(* CODESYS project functionresponse.library
   Company: KOSTAL GmbH & Co.KG
   DocFormat: reStructuredText
   DefaultNamespace: KOSTAL.AF2024.Core.functionResponse
   Version: 1.0.0.0
   Placeholder: KOSTAL.AF2024.Core.functionResponse
   Author: Frank Dümpelmann
   Title: KOSTAL.AF2024.Core.functionResponse

Project tree, tasks and I/O mapping:
  libraries: KOSTAL.AF2024.Core.Settings, * (KOSTAL GmbH & Co.KG); KOSTAL.AF2024.Core.System, * (KOSTAL GmbH & Co.KG)
  DUT/
    interface I_T_functionResponse: CopyTo, status, success
    interface I_T_functionResponse_CopyFrom: CopyFrom
    interface I_T_functionResponse_Owner: clear, CopyFrom, CopyTo, status, success
    function block T_functionResponse [ST]: clear, CopyFrom, CopyTo, status, success
  Project Information/
    function F_GetCompany [ST]
    function F_GetTitle [ST]
    function F_GetVersion [ST]
  Version/
    global variables Global_Version
*)

// Version/Global_Version
{attribute 'TcGenerated'}
{attribute 'no-analysis'}
{attribute 'linkalways'}
// This function has been automatically generated from the project information.
VAR_GLOBAL CONSTANT
	{attribute 'const_non_replaced'}
	stLibVersion_KOSTAL_AF2024_Core_functionResponse : ST_LibVersion := (iMajor := 1, iMinor := 0, iBuild := 0, iRevision := 0, nFlags := 0, sVersion := '1.0.0.0');
END_VAR

// DUT/I_T_functionResponse
INTERFACE I_T_functionResponse EXTENDS KOSTAL_AF2024_Core_System.I_Interface

METHOD PUBLIC CopyTo
VAR_INPUT
	IN : I_T_functionResponse_CopyFrom;
END_VAR
END_METHOD

PROPERTY PUBLIC status : KOSTAL_AF2024_Core_Settings.T_MaxString
GET
END_GET
END_PROPERTY

PROPERTY PUBLIC success : BOOL
GET
END_GET
END_PROPERTY

END_INTERFACE

// DUT/I_T_functionResponse_CopyFrom
INTERFACE I_T_functionResponse_CopyFrom EXTENDS KOSTAL_AF2024_Core_System.I_Interface

METHOD PUBLIC CopyFrom
VAR_INPUT
	IN	: I_T_functionResponse;
END_VAR
END_METHOD

END_INTERFACE

// DUT/I_T_functionResponse_Owner
INTERFACE I_T_functionResponse_Owner EXTENDS KOSTAL_AF2024_Core_System.I_Interface

METHOD PUBLIC clear
END_METHOD

METHOD PUBLIC CopyFrom
VAR_INPUT
	IN	: I_T_functionResponse;
END_VAR
END_METHOD

METHOD PUBLIC CopyTo
VAR_INPUT
	IN : I_T_functionResponse_CopyFrom;
END_VAR
END_METHOD

PROPERTY PUBLIC status : KOSTAL_AF2024_Core_Settings.T_MaxString
GET
END_GET
SET
END_SET
END_PROPERTY

PROPERTY PUBLIC success : BOOL
GET
END_GET
SET
END_SET
END_PROPERTY

END_INTERFACE

// DUT/T_functionResponse
(*

:Author: Frank Dümpelmann <f.duempelmann@kostal.com>
:Date: 2018-10-26

Function
========
Data type for function responses

Methods and Properties
======================
| success 	:BOOL 	Function or method sucessfully finished
| status	:STRING Fault description in case of failure
| clear()	METHOD	Reset all values	
*)
{attribute 'enable_dynamic_creation'}
FUNCTION_BLOCK PUBLIC T_functionResponse IMPLEMENTS I_T_functionResponse, I_T_functionResponse_CopyFrom, I_T_functionResponse_Owner

VAR
	_success	: BOOL;	//BOOL
	_status		: KOSTAL_AF2024_Core_Settings.T_MaxString;
END_VAR

METHOD PUBLIC clear

_status		:= "";
_success	:= FALSE;
END_METHOD

METHOD PUBLIC CopyFrom
VAR_INPUT
	IN	: I_T_functionResponse;
END_VAR

IF IN = 0 THEN RETURN;	END_IF

_success:= IN.success;
_status	:= IN.status;
END_METHOD

METHOD PUBLIC CopyTo
VAR_INPUT
	IN : I_T_functionResponse_CopyFrom;
END_VAR

IF IN = 0 THEN RETURN;	END_IF

IN.CopyFrom(THIS^);
END_METHOD

PROPERTY PUBLIC status : KOSTAL_AF2024_Core_Settings.T_MaxString
GET

status:= _status;
END_GET
SET

_status:= status;
END_SET
END_PROPERTY

PROPERTY PUBLIC success : BOOL
GET

success:= _success;
END_GET
SET

_success:= success;
END_SET
END_PROPERTY

END_FUNCTION_BLOCK

// Project Information/F_GetCompany
// This function has been automatically generated from the project information.
{attribute 'signature_flag' := '1073741824'}
{attribute 'TcGenerated'}
{attribute 'no-analysis'}
FUNCTION F_GetCompany : WSTRING
VAR_INPUT
	
END_VAR

F_GetCompany := "KOSTAL GmbH & Co.KG";

END_FUNCTION

// Project Information/F_GetTitle
// This function has been automatically generated from the project information.
{attribute 'signature_flag' := '1073741824'}
{attribute 'TcGenerated'}
{attribute 'no-analysis'}
FUNCTION F_GetTitle : WSTRING
VAR_INPUT
	
END_VAR

F_GetTitle := "KOSTAL.AF2024.Core.functionResponse";

END_FUNCTION

// Project Information/F_GetVersion
// This function has been automatically generated from the project information.
{attribute 'signature_flag' := '1073741824'}
{attribute 'TcGenerated'}
{attribute 'no-analysis'}
FUNCTION F_GetVersion : ST_LibVersion
VAR_INPUT
	
END_VAR

F_GetVersion.iMajor := 1;
F_GetVersion.iMinor := 0;
F_GetVersion.iBuild := 0;
F_GetVersion.iRevision := 0;
F_GetVersion.sVersion := '1.0.0.0';
F_GetVersion.nFlags := 0;

END_FUNCTION
